Fanuc KAREL source: KT00889.KL

PROGRAM KT00889
%NOLOCKGROUP
VAR
  P1: XYZWPR
  P2: XYZWPR
  OUT: POSITION
BEGIN
  P1.X = 1.0
  P2.Y = 2.0
  P1.X = 1.0
  P2.Y = 2.0
  OUT = INV(P1)
END KT00889
